FUNCTION_BLOCK DropConstraint
VAR_INPUT
	kDrop: DINT;
END_VAR
VAR_OUTPUT
END_VAR
VAR_IN_OUT
	iA: ARRAY[0..243] OF BOOL;
	nA: DINT;
	iC: ARRAY[0..243] OF DINT;
END_VAR
VAR
	i: DINT;
END_VAR



IF kDrop > 0 THEN 
    iA[iC[kDrop - 1] - 1] := FALSE;

    IF kDrop < nA THEN 
        i := kDrop;
        WHILE i <= (nA - 1) DO
            iC[i - 1] := iC[i];
            i := i + 1;
        END_WHILE;
    END_IF;

    iC[nA - 1] := 0;
    nA := nA - 1;
END_IF;

END_FUNCTION_BLOCK

(* stored: Version 1.1.0.1, ProductVersion 3.1.4024.9
   POU DropConstraint: Id {43ab0fed-5f30-46c2-9f92-2ccd622d101b}, SpecialFunc None *)
